// TIA Portal V20 export
// export: Created 2026-10-20T12:39:40.4550332Z, ExportSetting WithDefaults, DisplayName Totally Integrated Automation Portal, DisplayVersion V20 Update 6, DisplayName TIA Portal Openness, DisplayVersion V20 Update 6, DisplayName TIA Portal Version Control Interface, DisplayVersion V20 Update 6, DisplayName SINAMICS Startdrive Advanced, DisplayVersion V20 SP1, DisplayName SINAMICS Startdrive G130, G150, S120, S150, SINAMICS MV, G220, S200, S210, DisplayVersion V20 SP1, DisplayName SINAMICS Startdrive G110M, G120, G120C, G120D, G120P, G115D, DisplayVersion V20 SP1, DisplayName STEP 7 Professional, DisplayVersion V20 Update 6, DisplayName STEP 7 Safety, DisplayVersion V20 Update 2, DisplayName WinCC Basic/Comfort/Advanced, DisplayVersion V20 Update 6, DisplayName WinCC Unified, DisplayVersion V20 Update 6
DATA_BLOCK "Bypass"   // DB9
{ S7_Optimized_Access := 'TRUE' }
VERSION : 0.1
// stored: AutoNumber true, DBAccessibleFromOPCUA true, IsOnlyStoredInLoadMemory false, IsRetainMemResEnabled false, IsWriteProtectedInAS false, MemoryReserve 100
   VAR RETAIN
      Main_Panel { S7_SetPoint := 'True'} : "Safety_Bypass_MainPanel";
      Remote_Panel_1 : "Safety_Bypass_RemotePanel";
      Remote_Panel_2 { S7_SetPoint := 'True'} : "Safety_Bypass_RemotePanel";
      Remote_Panel_3 { S7_SetPoint := 'True'} : "Safety_Bypass_RemotePanel";
      Remote_Panel_4 { S7_SetPoint := 'True'} : "Safety_Bypass_RemotePanel";
      Remote_Panel_5 { S7_SetPoint := 'True'} : "Safety_Bypass_RemotePanel";
   END_VAR
BEGIN
   Main_Panel.Estop_Cabinet := FALSE;
END_DATA_BLOCK
